// SIMATIC S7-200 project (STEP 7-Micro/WIN), CPU 226 CN REL 02.01

SYMBOL_TABLE ????1
boton_sb1        I2.5
boton_sb2        I2.4
selector         I2.7
parada           I2.6
act1             Q0.0
act2             Q0.1
act3             Q0.3
act4             Q0.4
act5             Q0.5
act6             Q0.6
act7             Q0.7
act8             Q1.0
END_SYMBOL_TABLE

ORGANIZATION_BLOCK ???:OB1
TITLE=????
BEGIN
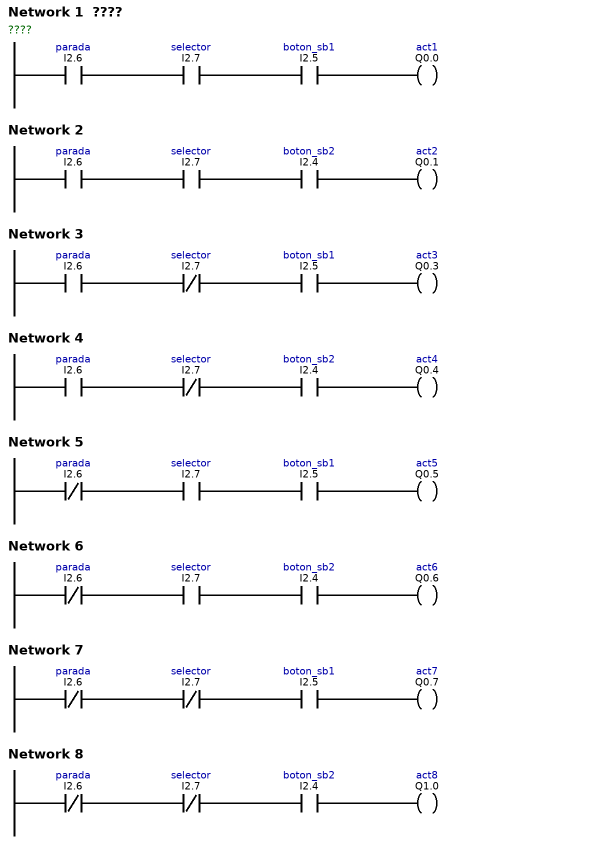
Network 1 // ????
// ????
LD     parada:I2.6
A      selector:I2.7
A      boton_sb1:I2.5
=      act1:Q0.0
Network 2
LD     parada:I2.6
A      selector:I2.7
A      boton_sb2:I2.4
=      act2:Q0.1
Network 3
LD     parada:I2.6
AN     selector:I2.7
A      boton_sb1:I2.5
=      act3:Q0.3
Network 4
LD     parada:I2.6
AN     selector:I2.7
A      boton_sb2:I2.4
=      act4:Q0.4
Network 5
LDN    parada:I2.6
A      selector:I2.7
A      boton_sb1:I2.5
=      act5:Q0.5
Network 6
LDN    parada:I2.6
A      selector:I2.7
A      boton_sb2:I2.4
=      act6:Q0.6
Network 7
LDN    parada:I2.6
AN     selector:I2.7
A      boton_sb1:I2.5
=      act7:Q0.7
Network 8
LDN    parada:I2.6
AN     selector:I2.7
A      boton_sb2:I2.4
=      act8:Q1.0
END_ORGANIZATION_BLOCK
